Staubli VAL3: showCoord.pgx

program showCoord(num x_nIndex)
begin
  sTRSF[0]=toString(".2",safeTemp:sSPoint[x_nIndex].pPointRx.trsf.x)
  sTRSF[1]=toString(".2",safeTemp:sSPoint[x_nIndex].pPointRx.trsf.y)
  sTRSF[2]=toString(".2",safeTemp:sSPoint[x_nIndex].pPointRx.trsf.z)
  sTRSF[3]=toString(".2",safeTemp:sSPoint[x_nIndex].pPointRx.trsf.rx)
  sTRSF[4]=toString(".2",safeTemp:sSPoint[x_nIndex].pPointRx.trsf.ry)
  sTRSF[5]=toString(".2",safeTemp:sSPoint[x_nIndex].pPointRx.trsf.rz)
end
